(* IEC 61131-3 sources: OpenPlc_Lezioni/sfdb_led/build, 2 files *)

(* ---- plc.st ---- *)
TYPE
  LOGLEVEL : (CRITICAL, WARNING, INFO, DEBUG) := INFO;
END_TYPE

FUNCTION_BLOCK LOGGER
  VAR_INPUT
    TRIG : BOOL;
    MSG : STRING;
    LEVEL : LOGLEVEL := INFO;
  END_VAR
  VAR
    TRIG0 : BOOL;
  END_VAR

  IF TRIG AND NOT TRIG0 THEN
  {{
   LogMessage(GetFbVar(LEVEL),(char*)GetFbVar(MSG, .body),GetFbVar(MSG, .len));
  }}
  END_IF;
  TRIG0:=TRIG;
END_FUNCTION_BLOCK

PROGRAM program0
  VAR
    bt1 : BOOL;
    led_verde : BOOL;
    T1 : BOOL;
    SR0 : SR;
    TON0 : TON;
  END_VAR

  SR0(S1 := bt1, R := T1);
  led_verde := SR0.Q1;
  TON0(IN := SR0.Q1, PT := T#10s);
  T1 := TON0.Q;
END_PROGRAM

CONFIGURATION Config0

  RESOURCE Res0 ON PLC
    TASK task0(INTERVAL := T#20ms,PRIORITY := 0);
    PROGRAM instance0 WITH task0 : program0;
  END_RESOURCE
END_CONFIGURATION

(* ---- generated_plc.st ---- *)
PROGRAM program0
  VAR
    bt1 : BOOL;
    led_verde : BOOL;
    T1 : BOOL;
    SR0 : SR;
    TON0 : TON;
  END_VAR

  SR0(S1 := bt1, R := T1);
  led_verde := SR0.Q1;
  TON0(IN := SR0.Q1, PT := T#10s);
  T1 := TON0.Q;
END_PROGRAM

CONFIGURATION Config0

  RESOURCE Res0 ON PLC
    TASK task0(INTERVAL := T#20ms,PRIORITY := 0);
    PROGRAM instance0 WITH task0 : program0;
  END_RESOURCE
END_CONFIGURATION
